TYPE ST_ROBOTTOPLC :
STRUCT
	arbyInput				:ARRAY[0..63] OF BYTE;
END_STRUCT
END_TYPE

(* stored: Version 1.1.0.1, ProductVersion 3.1.4024.15
   DUT ST_ROBOTTOPLC: Id {037e5b95-2935-4edd-8fd2-9eb71b3bb654} *)
